(* IEC 61131-3 sources: ATCMcontrol_Engineering/src/COM/softing/fc/AddOns/Softing/4CPCTarget/Libs/ATCM_Communication, 12 files *)

(* ---- CONNECT.ST ---- *)
(*[[
    UserURL= "ATCM:CONNECT.htm"
]]*)

(* Communication Function Blocks, see IEC 1131-5
 * Implements the CONNECT communication function block
 *
*)

FUNCTION_BLOCK CONNECT      (* Connection management *)
VAR_INPUT
	EN_C    : BOOL := FALSE;   (* enable/startup connection *)
	PARTNER : COMM_PARTNER;    (* identifies communication partner and comm. deployment *)
END_VAR
VAR_OUTPUT
	VALID  : BOOL := FALSE;    (* connection is valid/established *)
	ERROR  : BOOL := FALSE;    (* new non-zero STATUS received *)
    STATUS : DINT := CFB_NoError;   (* last detected status *)
	ID     : COMM_CHANNEL;     (* established communication channel *)
END_VAR

VAR
    iType       : DINT;
    hChannel    : DINT;
    sParam      : WSTRING;
    bError   : BOOL;            (* true if error occured *)
    iNewStatus : DINT;          (* new status *)
    iFbState : DINT := 0;       (* state of function block:*)
                                (*  0: INIT
                                    1: IDLE
                                    2: CONNECTING
                                    3: CHECKING
                                    4: CONNECTED
                                    5: CLOSING
                                    6: CONCLUDING
                                    7: RETRY
                                    8: ABORT
                                    10: ERROR
                                *)
END_VAR

VAR_NATIVE
    static CommFBFactory g_commFBFact = new CommFBFactory();
    private CommFB comm = null;
    private int hChannel;
    private int iType;
    public void release()
    {
        if (comm != null)
        {
            CommFBFactory.removeCommFB(hChannel, iType);
            comm.closeConn();
            comm.release();
            comm = null;
        }
        super.release();
    }
END_VAR

VAR_NATIVE#movetop
import COM.softing.fc.CC.commFB.*;
END_VAR

(*
NATIVE
END_VAR
*)

(* Init local variables *)
hChannel := ID.hChannel;
iType := ID.iCommType;
bError := FALSE;
iNewStatus := CFB_NoError;

(* Init OutVars *)
ERROR := FALSE;

(* INIT funciton Block *)
IF iFbState = 0 THEN
    VALID := FALSE;
    STATUS := CFB_NoError;

    (* fast initialization => next fb state: idle *)
    iFbState := 1;
END_IF;

(* IDLE until new connect request *)
IF iFbState = 1 THEN
    IF EN_C THEN
        VALID := FALSE;
        ID.hChannel := -1;  (* not valid *)
        hChannel := -1;

        iType := PARTNER.iCommType;
        sParam := PARTNER.sParam;
        ID.iCommType := iType;
        ID.iTimeout := PARTNER.iTimeout;
        (* next state connecting *)
        iFbState := 2;
    ELSE
        (* Idle...*)
        RETURN;
    END_IF;
END_IF;

(* CONNECTING *)
IF iFbState = 2 THEN
    IF EN_C THEN
        (* Open connection *)
        NATIVE
        //if there is an old commFB, KILL IT NOW!
        if (comm != null)
        {
            CommFBFactory.removeCommFB(hChannel, iType);
            comm.closeConn();
            comm.release();
            comm = null;
        }
        // create new CommFB
        comm = CommFBFactory.createCommFB(iType = _itype.getInt());
        if (comm == null)
        {
            _berror.putBool(true);
            _inewstatus.putInt(-4); // CFB_ErrOutOfMemory
        }
        else
        {
            // open connection
            if (comm.openConn(_sparam.getString()))
            {
                hChannel = CommFBFactory.addCommFBToMap(comm);
                _hchannel.putInt(hChannel);
            }
            else
            {
                _berror.putBool(true);
                _inewstatus.putInt(comm.getConnStatus()); // CFB_...
                comm = null;
            }
        }
        END_NATIVE;

        IF bError THEN
            (* next state error *)
            iFbState := 10;
            GOTO error;
        ELSE
            (* next state checking *)
            iFbState := 3;
        END_IF;

    ELSE (* EN_C = FALSE *)
        (* Abort => next state idle *)
        iFbState := 1;
        RETURN;
    END_IF;
END_IF;

(* CHECKING *)
IF iFbState = 3 THEN
    NATIVE
    if (comm == null)
    {
        _berror.putBool(true);
        _inewstatus.putInt(7);  // CFB_ErrRemoteWrongState
        // next state error
        _ifbstate.putInt(10);
    }
    else if (!comm.checkConn())
    {
        _berror.putBool(true);
        _inewstatus.putInt(1);  // CFB_ErrLowLayer
        // next state abort
        _ifbstate.putInt(8);
    }
    END_NATIVE;

    IF bError = FALSE THEN
        ID.hChannel := hChannel;
        VALID := TRUE;
        (* next state connected *)
        iFbState := 4;
        (* wait for next cycle... *)
        RETURN;
    END_IF;
END_IF;

(* CONNECTED *)
IF iFbState = 4 THEN
    IF EN_C = FALSE THEN
        (* next state closing *)
        iFbState := 5;
    ELSE
        NATIVE
        if (comm == null)
            _berror.putBool(true);
        END_NATIVE;

        IF bError THEN
            iNewStatus := CFB_ErrRemoteWrongState;
            (* next state error *)
            iFbState := 10;
            GOTO error;
        ELSE
            (* check if connection is closed by the remote station *)
            NATIVE
            if (comm.isRemoteClosing())
            {
                // next state concluding
                _ifbstate.putInt(6);
                // wait for next cycle...
                return;
            }
            END_NATIVE;

            (* check if connection is still alive *)
            NATIVE
            if (!comm.checkConn())
            {
                _berror.putBool(true);
                _inewstatus.putInt(1); // CFB_ErrLowLayer
                // next state retry
                _ifbstate.putInt(7);
            }
            END_NATIVE;
        END_IF;
    END_IF;
END_IF;

(* CLOSING *)
IF iFbState = 5 THEN
    NATIVE
    if (comm != null)
    {
        CommFBFactory.removeCommFB(hChannel, iType);
        comm.closeConn();
        comm.release();
        comm = null;
    }
    END_NATIVE;

    VALID := FALSE;
    ID.hChannel := -1;
    (* next state idle *)
    iFbState := 1;
END_IF;

(* CONCLUDING *)
IF iFbState = 6 THEN
    NATIVE
    if (comm != null)
    {
        CommFBFactory.removeCommFB(hChannel, iType);
        comm.closeConn();
        comm.release();
        comm = null;
    }
    END_NATIVE;

    VALID := FALSE;
    ID.hChannel := -1;
    STATUS := CFB_ErrResetReceived;
    (* next state idle *)
    iFbState := 1;
END_IF;

(* RETRY *)
IF iFbState = 7 THEN
    NATIVE
    if (comm != null)
    {
        CommFBFactory.removeCommFB(hChannel, iType);
        comm.closeConn();
        comm.release();
        comm = null;
    }
    END_NATIVE;
    (* next state error *)
    iFbState := 10;
    GOTO error;
END_IF;

(* ABORT *)
IF iFbState = 8 THEN
    NATIVE
    if (comm != null)
    {
        CommFBFactory.removeCommFB(hChannel, iType);
        comm.closeConn();
        comm.release();
        comm = null;
    }
    END_NATIVE;
    (* next state error *)
    iFbState := 10;
    GOTO error;
END_IF;

(* ERROR *)
error:
IF iFbState = 10 THEN
    NATIVE
    if (comm != null)
    {
        CommFBFactory.removeCommFB(hChannel, iType);
        comm.closeConn();
        comm.release();
        comm = null;
    }
    END_NATIVE;

    VALID := FALSE;
    ERROR := TRUE;
    STATUS := iNewStatus;

    iFbState := 1;
    RETURN;
END_IF;

END_FUNCTION_BLOCK

(* ---- RCV.ST ---- *)
(*[[
]]*)

(* Communication Function Blocks, see IEC 1131-5
 * Implements the RCV communication function block
 *
*)

NATIVE
import COM.softing.fc.CC.commFB.*;
END_NATIVE

FUNCTION_BLOCK RCV      (* Interlocked control, responder*)
VAR_INPUT
    EN_R   : BOOL;          (* Enable to receive data *)
    RESP   : BOOL (*R_EDGE*);   (* Request to send response data *)
    ID     : COMM_CHANNEL;  (* Communication channel *)
    R_ID   : WSTRING;       (* Remote function block *)
    EXPECT : DINT;          (* non-IEC: number of bytes to receive *)
(*    SD_1   : ANY;*)           (* User data to send *)
(*    SD_m   : ANY; *)
END_VAR

VAR_OUTPUT
NDR    : BOOL;              (* New user data received *)
ERROR  : BOOL;              (* New non-zero STATUS received *)
STATUS : DINT;              (* Last detected status *)

RD_1   : WSTRING; (*ANY*)       (* Received user data *)
(*RD_n   : ANY;*)         (*  It is not required that m=n *)
END_VAR                 (*  either m, n, or both may be 0*)

    (* is not implemented yet !! *)
    ERROR := TRUE;
    STATUS := CFB_ErrNotImpl;

NATIVE
END_NATIVE;

END_FUNCTION_BLOCK

(* ---- SEND.ST ---- *)
(*[[
]]*)

(* Communication Function Blocks, see IEC 1131-5
 * Implements the SEND communication function block
 *
*)

NATIVE
import COM.softing.fc.CC.commFB.*;
END_NATIVE

FUNCTION_BLOCK SEND     (* Interlocked control, requester*)
VAR_INPUT
    REQ    : BOOL (*R_EDGE*);       (* Request to send with raising edge*)
    R      : BOOL (*R_EDGE*);       (* Reset local, remote function *)
    ID     : COMM_CHANNEL;      (* Communication channel *)
    R_ID   : WSTRING;           (* Remote function block *)
    SD_1   : WSTRING;  (*ANY*)  (* User data to send *)
END_VAR

VAR_OUTPUT
    NDR    : BOOL;          (* New user data received *)
    ERROR  : BOOL;        (* New non-zero STATUS received *)
    STATUS : DINT;        (* Last detected status *)
(*    RD_1   : ANY;*)         (* Received user data *)
END_VAR                 (*   either m, n, or both may be 0*)

    (* is not implemented yet !! *)
    ERROR := TRUE;
    STATUS := CFB_ErrNotImpl;

NATIVE
END_NATIVE;

END_FUNCTION_BLOCK

(* ---- SER_READ.ST ---- *)
(*[[
    UserURL= "ATCM:SER_READ.htm"
]]*)

(* Communication Function Blocks, see IEC 1131-5 for serial communication
 * Derived from the READ communication function block
 * differs in RD_LEN1, resp. RD_1 from READ in IEC 1131-5!
*)

FUNCTION_BLOCK SER_READ     (* Polled data acquisition *)
VAR_INPUT
    REQ      : BOOL R_EDGE := FALSE;    (* Request *)
    ID       : COMM_CHANNEL;    (* Communication channel *)
    RD_LEN_1 : DINT;            (* Min. length of the data to be received *)
    READ_ALL : BOOL := FALSE;   (* TRUE: all available data will be read, at least RD_LEN_1 *)
END_VAR

VAR_OUTPUT
    NDR    : BOOL;              (* New user data received *)
    ERROR  : BOOL;              (* New non-zero STATUS received *)
    STATUS : DINT;              (* Last detected status *)
    RD_1   : BYTE_STRING;       (* Received user data *)
END_VAR

VAR
    hChannel : DINT;
    iType    : DINT;
    bError   : BOOL;            (* true if error occured *)
    iNewStatus : DINT;          (* new status *)
    iFbState : DINT := 0;       (* state of function block:*)
                                (*  0: INIT
                                    1: IDLE
                                    2: WAITING
                                    3: CHECKING
                                    4: HAVE_DATA
                                    10: ERROR
                                *)
    timer    : TON;             (* timer for read timeout *)
    timer_IN : BOOL;
    timer_PT : TIME;
    bTimeout : BOOL;
END_VAR

VAR_NATIVE
    private CommFB comm;
END_VAR
VAR_NATIVE#movetop
import COM.softing.fc.CC.commFB.*;
import COM.softing.fc.CC.utility.*;
END_VAR

(* Init local variables*)
hChannel := ID.hChannel;
iType := ID.iCommType;
bError := FALSE;

(* Init OutVars *)
NDR := FALSE;
ERROR := FALSE;

(* INIT funciton Block *)
IF iFbState = 0 THEN
    STATUS := CFB_NoError;

    (* fast initialization => goto next state IDLE*)
    iFbState := 1;
END_IF;

(* get CommFB *)
NATIVE
    comm = CommFBFactory.lookUpCommFB(_hchannel.getInt(), _itype.getInt());
    if (comm == null)
    {
        _berror.putBool(true);
    }
END_NATIVE;
IF bError THEN
    iNewStatus := CFB_ErrInvalidCommChannel;
    iFbState := 10;
    GOTO error;
END_IF;

(* IDLE until new read request at raising edge of REQ input *)
IF iFbState = 1 THEN
    IF REQ THEN
        NATIVE
        // check if read is not active
        synchronized(comm) {
          if (comm.isReadActive())
            _berror.putBool(true);
          else
            comm.setReadActive(true);
        }
        END_NATIVE;

        IF bError THEN
            iNewStatus := CFB_ErrRemoteWrongState;
            iFbState := 10;
            GOTO error;
        END_IF;
        (* Start read request asynchronously *)
        (* reset timer *)
        bTimeout := FALSE;
        timer_IN := FALSE;
        timer_PT := DINT_TO_TIME(ID.iTimeout);
        timer(IN := timer_IN, PT := timer_PT);

        NATIVE
        // start read request
        if (!comm.readAsync(_rd_len_1, _read_all, (ByteString)_rd_1))
        {
            _berror.putBool(true);
            _inewstatus.putInt(comm.getReadStatus()); // CFB_...
            comm.setReadActive(false);
        }
        END_NATIVE;

        IF bError THEN
            iFBState := 10;
            GOTO error;
        END_IF;

        (* init new timer *)
        IF ID.iTimeout > 0 THEN
            timer_IN := TRUE;
        ELSE
            timer_IN := FALSE;
        END_IF;

        (* Next state WAITING *)
        iFbState := 2;

    ELSE
        (* Idle...*)
        RETURN;
    END_IF;
END_IF;

(* WAITING: wait for completion *)
IF iFbState = 2 THEN
    (* refresh timer *)
    timer(IN := timer_IN, PT := timer_PT);
    bTimeout := timer.Q;

    (* Wait for data *)
    NATIVE
    if (comm.hasReadCompleted())
    {
        // check status if error occured
        int iStat = comm.getReadStatus();
        if (iStat == 0)
        {
            // read finished : next state CHECKING
            _inewstatus.putInt(0);
            _ifbstate.putInt(3);
        }
        else
        {
            // error!
            _berror.putBool(true);
            _inewstatus.putInt(iStat); // CFB_...
            comm.setReadActive(false);
        }
    }
    else
    {
        // request pending!
        if (_btimeout.getBool())
        {
            // cancel read request
            comm.cancelReadRequest();
            _berror.putBool(true);
            comm.setReadActive(false);
        }
        else
        {
            // wait for next cycle...
            return;
        }
    }
    END_NATIVE;
    IF bError THEN
        IF bTimeout THEN
            iNewStatus := CFB_ErrTimeout;
        ELSE
            ; (* iNewStatus already set *)
        END_IF;
        iFBState := 10;
        GOTO error;
    END_IF;

END_IF;

(* CHECKING data type match *)
IF iFbState = 3 THEN
    NATIVE
    if (!comm.verifyData())
    {
        _berror.putBool(true);
        comm.setReadActive(false);
    }
    END_NATIVE;
    IF bError THEN
        iNewStatus := CFB_ErrTypeMismatch;
        iFBState := 10;
        GOTO error;
    ELSE
        (* next state: HAVE DATA *)
        iFBState := 4;
    END_IF;
END_IF;

(* HAVE DATA *)
IF iFbState = 4 THEN
    (* copy data to RD_1 *)
    NATIVE
    comm.depositData();
    comm.setReadActive(false);
    END_NATIVE;

    NDR := TRUE;
    ERROR := FALSE;
    STATUS := 0;

    (* next state: IDLE *)
    iFbState := 1;
    RETURN;
END_IF;

(* ERROR *)
error:
IF iFbState = 10 THEN
    NDR := FALSE;
    ERROR := TRUE;
    STATUS := iNewStatus;

    iFbState := 1;
    RETURN;
END_IF;

END_FUNCTION_BLOCK

(* ---- SER_WRITE.st ---- *)
(*[[
    UserURL= "ATCM:SER_WRITE.htm"
]]*)

(* Communication Function Blocks, see IEC 1131-5 for serial communication
 * Derived from the WRITE communication function block
 * differs in SD_1 from WRITE in IEC 1131-5!
*)

FUNCTION_BLOCK SER_WRITE            (* Parametric control *)
VAR_INPUT
    REQ    : BOOL R_EDGE := FALSE;  (* Request *)
    ID     : COMM_CHANNEL;          (* Communication channel *)
    SD_1   : BYTE_STRING ;          (* value of to be set *)
END_VAR

VAR_OUTPUT
    DONE   : BOOL;        (* Function performed *)
    ERROR  : BOOL;        (* New non-zero STATUS received *)
    STATUS : DINT;        (* Last detected status *)
END_VAR

VAR
    hChannel : DINT;
    iType    : DINT;
    bError   : BOOL;            (* true if error occured *)
    iNewStatus : DINT;          (* new status *)
    iFbState : DINT := 0;       (* state of function block:*)
                                (*  0: INIT
                                    1: IDLE
                                    2: WAITING
                                    4: HAVE_IT
                                    10: ERROR
                                *)
    timer    : TON;             (* timer for write timeout *)
    timer_IN : BOOL;
    timer_PT : TIME;
    bTimeout : BOOL;
END_VAR

VAR_NATIVE
    private CommFB comm;
END_VAR
VAR_NATIVE#movetop
import COM.softing.fc.CC.commFB.*;
import COM.softing.fc.CC.utility.*;
END_VAR

(* INIT local variables*)
hChannel := ID.hChannel;
iType := ID.iCommType;
bError := FALSE;

(* Init OutVars *)
DONE := FALSE;
ERROR := FALSE;

(* Init funciton Block *)
IF iFbState = 0 THEN
    STATUS := CFB_NoError;

    (* fast initialization => goto state IDLE *)
    iFbState := 1;
END_IF;

(* get CommFB *)
NATIVE
    comm = CommFBFactory.lookUpCommFB(_hchannel.getInt(), _itype.getInt());
    if (comm == null)
    {
        _berror.putBool(true);
    }
END_NATIVE;
IF bError THEN
    iNewStatus := CFB_ErrInvalidCommChannel;
    iFbState := 10;
    GOTO error;
END_IF;

(* IDLE until new write request at raising edge of REQ input *)
IF iFbState = 1 THEN
    IF REQ THEN
        NATIVE
        // check if write is not active
        synchronized(comm) {
          if (comm.isWriteActive())
            _berror.putBool(true);
          else
            comm.setWriteActive(true);
        }
        END_NATIVE;

        IF bError THEN
            iNewStatus := CFB_ErrRemoteWrongState;
            iFbState := 10;
            GOTO error;
        END_IF;

        (* Start write request asynchronously *)
        (* reset timer *)
        bTimeout := FALSE;
        timer_IN := FALSE;
        timer_PT := DINT_TO_TIME(ID.iTimeout);
        timer(IN := timer_IN, PT := timer_PT);

        NATIVE
        // source: locVars[2])
        if (!comm.writeAsync((ByteString)_sd_1))
        {
            _berror.putBool(true);
            _inewstatus.putInt(comm.getWriteStatus()); // CFB_...
            comm.setWriteActive(false);
        }
        END_NATIVE;

        IF bError THEN
            iFBState := 10;
            GOTO error;
        END_IF;

        (* init new timer *)
        IF ID.iTimeout > 0 THEN
            timer_IN := TRUE;
        ELSE
            timer_IN := FALSE;
        END_IF;

        (* Sext state WAITING *)
        iFbState := 2;

    ELSE
        (* Idle...*)
        RETURN;
    END_IF;
END_IF;

(* WAITING: wait for completion *)
IF iFbState = 2 THEN
    (* refresh timer *)
    timer(IN := timer_IN, PT := timer_PT);
    bTimeout := timer.Q;

    (* Wait for completion *)
    NATIVE
    if (comm.hasWriteCompleted())
    {
        // check status if error occured
        int iStat = comm.getWriteStatus();
        if (iStat == 0)
        {
            // write finished: next state HAVE IT
            _inewstatus.putInt(0);
            _ifbstate.putInt(4);
        }
        else
        {
            // error!
            _berror.putBool(true);
            _inewstatus.putInt(iStat); // CFB_...
            comm.setWriteActive(false);
        }
    }
    else
    {
        // request pending!
        if (_btimeout.getBool())
        {
            // cancel write request
            comm.cancelWriteRequest();
            _berror.putBool(true);
            comm.setWriteActive(false);
        }
        else
        {
            // wait for next cycle...
            return;
        }
    }
    END_NATIVE;
    IF bError THEN
        IF bTimeout THEN
            iNewStatus := CFB_ErrTimeout;
        ELSE
            ; (* iNewStatus already set *)
        END_IF;
        iFBState := 10;
        GOTO error;
    END_IF;

END_IF;

(* HAVE IT *)
IF iFbState = 4 THEN
    NATIVE
    comm.setWriteActive(false);
    END_NATIVE;
    DONE := TRUE;
    ERROR := FALSE;
    STATUS := 0;

    iFbState := 1;
    RETURN;
END_IF;

(* ERROR *)
error:
IF iFbState = 10 THEN
    DONE := FALSE;
    ERROR := TRUE;
    STATUS := iNewStatus;

    iFbState := 1;
    RETURN;
END_IF;

END_FUNCTION_BLOCK

(* ---- STATUS.ST ---- *)
(*[[
]]*)

(* Communication Function Blocks, see IEC 1131-5
 * Implements the STATUS communication function block
 *
*)

NATIVE
import COM.softing.fc.CC.commFB.*;
END_NATIVE

FUNCTION_BLOCK STATUS   (* Device verification - requester *)
VAR_INPUT
    REQ    : BOOL (*R_EDGE*);   (* Request *)
    ID     : COMM_CHANNEL;  (* Communication channel *)
END_VAR

VAR_OUTPUT
    NDR    : BOOL;        (* New user data received *)
    ERROR  : BOOL;        (* New non-zero STATUS received *)
    STATUS : DINT;        (* Last detected status *)
    PHYS   : DINT;        (* Physical status of remote *)
                          (*   communication partner   *)
    LOG    : DINT;        (* Logical status of remote *)
                          (*   communication partner   *)
    LOCAL  : ARRAY[0..7] OF WORD;  (* Local status of remote *)
END_VAR

    (* is not implemented yet !! *)
    ERROR := TRUE;
    STATUS := CFB_ErrNotImpl;
NATIVE
END_NATIVE;

END_FUNCTION_BLOCK

(* ---- UDP_CONNECT.st ---- *)
(*[[
    UserURL= "ATCM:UDP_CONNECT.htm"
]]*)

(*
 *  UDP datagram communication Function Blocks
 *  UDP_CONNECT allows to open and close a socket
 *  this FunctionBlock should be called only once, when the
 *  socket should be opened or closed
 *)

FUNCTION_BLOCK UDP_CONNECT

VAR_INPUT
    EN_C : BOOL;           (* true: open and connect the socket *)
                           (*   the field LocalPort of SOCKET_HANDLE has to be filled
                                with the local port number where the socket wants to
                                receive messages *)
                           (* false: close the socket *)
                           (* this FunctionBlock should be called only once, when the
                              socket should be opened or closed *)
END_VAR

VAR_IN_OUT
    SOCKET_HANDLE : UDP_SOCKET_HANDLE;  (* a structure that describes the socket *)
END_VAR

VAR_OUTPUT
    VALID        : BOOL;   (* shows if the socket is open or close *)
    ERROR        : BOOL;   (* error information *)
    ERROR_NR     : DINT;
    ERROR_STRING : WSTRING;
END_VAR

VAR
    portNr : DInt;
    bc     : BOOL;
END_VAR

VAR_NATIVE#movetop
    import COM.softing.fc.CC.commFB.*;
END_VAR

if EN_C then
    portNr := SOCKET_HANDLE.localPort;
    bc := SOCKET_HANDLE.broadcastSocket;
    native
        ((COM.softing.fc.CC.commFB.UDPSocketHandle)_socket_handle).open(
                                    _portnr.getInt(),
                                    _bc.getBool(),
                                    _error,
                                    _error_nr,
                                    _error_string);
    end_native;
    VALID := not Error;
else
    native
        ((COM.softing.fc.CC.commFB.UDPSocketHandle)_socket_handle).close(
                                    _error,
                                    _error_nr,
                                    _error_string);
    end_native;
    VALID := false;
end_if;
;
END_FUNCTION_BLOCK

(* ---- UDP_LOOKUP.st ---- *)
(*[[
    UserURL= "ATCM:UDP_LOOKUP.htm"
]]*)

(*
 *  UDP datagram communication Function Blocks
 *  UDP_LOOKUP looks up the ip-address (abc.def.ghi.jkl)
 *  for a hostname, this has to be used in UDP_USEND
 *  UDP_LOOKUP works asynchron because lookup can take a while
 *)

FUNCTION_BLOCK UDP_LOOKUP

VAR_INPUT
    EN_L          : Bool;               (* if ENABLE_Lookup = true, do lookup else
                                            do nothing *)
    HOST_NAME     : WString;            (* the name of the host to look up *)
END_VAR

VAR_IN_OUT
    SOCKET_HANDLE : UDP_SOCKET_HANDLE;  (* a handle to a opened socket *)
END_VAR

VAR_OUTPUT
    READY         : Bool;               (* shows that the lookup thread has finished *)
    HOST_ADDRESS  : WString;            (* if the lookup succeeded, the address of the host *)
    ERROR         : Bool;               (* error information if an error happened *)
    ERROR_NR      : DInt;
    ERROR_STRING  : WString;
END_VAR

VAR_NATIVE#movetop
    import COM.softing.fc.CC.commFB.*;
END_VAR

native
    ((COM.softing.fc.CC.commFB.UDPSocketHandle)_socket_handle).lookup(
                                    _en_l.getBool(),
                                    _host_name.getString(),
                                    _ready,
                                    _host_address,
                                    _error,
                                    _error_nr,
                                    _error_string);
end_native;

;
END_FUNCTION_BLOCK

(* ---- UDP_URCV.st ---- *)
(*[[
    UserURL= "ATCM:UDP_URCV.htm"
]]*)

(*
 *  UDP datagram communication Function Blocks
 *  UDP_URCV allows to receive a message from a partner
 *  through an open socket, URCV looks if there is a new msg
 *  available. If yes it returns the msg data, else NDR shows
 *  that no new msg is available
 *)

FUNCTION_BLOCK UDP_URCV

VAR_INPUT
    EN_R     : BOOL;            (* true: look for a new msg, false: do nothing *)
    DATA_LEN : DINT;            (* the maximum number of bytes that want to be received *)
                                (*  udp is a datagram based protocol, that means the
                                    data will be received in packets. If the available packet is
                                    longer than DATA_LEN, only DATA_LEN bytes will be returend,
                                    the rest is lost *)
END_VAR

VAR_IN_OUT
    SOCKET_HANDLE : UDP_SOCKET_HANDLE;  (* a structure that describes the socket *)
END_VAR

VAR_OUTPUT
    RD_1         : BYTE_STRING;  (* contains the msg data, if a new msg has been received *)
    PARTNER_ADDR : WSTRING;      (* the address and port of the communication partner *)
    PARTNER_PORT : DINT;         (*    that sent the received msg *)
    NDR          : BOOL;         (* shows if a new msg has been received *)
    ERROR        : BOOL;         (* error information *)
    ERROR_NR     : DINT;
    ERROR_STRING : WSTRING;
END_VAR

VAR_NATIVE#movetop
    import COM.softing.fc.CC.commFB.*;
END_VAR

if (EN_R) then
    native
        ((COM.softing.fc.CC.commFB.UDPSocketHandle)_socket_handle).receive(
                _data_len.getInt(),
                _rd_1,
                _partner_addr,
                _partner_port,
                _error,
                _error_nr,
                _error_string);
    end_native;
    if (RD_1.size>0) then
        NDR := true;
    else
        NDR := false;
    end_if;
end_if;
;
END_FUNCTION_BLOCK

(* ---- UDP_USEND.st ---- *)
(*[[
    UserURL= "ATCM:UDP_USEND.htm"
]]*)

(*
 *  UDP datagram communication Function Blocks
 *  UDP_USEND allows to send a message to a partner
 *  through an open socket
 *)

FUNCTION_BLOCK UDP_USEND

VAR_INPUT
    REQ          : BOOL;             (* true: send the msg, false: do nothing *)
    PARTNER_ADDR : WSTRING;          (* the host address of the communication partner *)
    PARTNER_PORT : DINT;             (* the port number where the comm. partner receives its msgs *)
    SD_1         : BYTE_STRING;      (* the data of the msg that will be sent *)
END_VAR

VAR_IN_OUT
    SOCKET_HANDLE : UDP_SOCKET_HANDLE; (* a structure that describes the socket *)
END_VAR

VAR_OUTPUT
    ERROR        : BOOL;             (* error information *)
    ERROR_NR     : DINT;
    ERROR_STRING : WSTRING;
END_VAR

VAR_NATIVE#movetop
    import COM.softing.fc.CC.commFB.*;
END_VAR

if (REQ) then
    native
        ((COM.softing.fc.CC.commFB.UDPSocketHandle)_socket_handle).send(
            _partner_addr.getString(),
            _partner_port.getInt(),
            _sd_1,
            _error,
            _error_nr,
            _error_string);
    end_native;
end_if;

END_FUNCTION_BLOCK

(* ---- USTATUS.ST ---- *)
(*[[
]]*)

(* Communication Function Blocks, see IEC 1131-5
 * Implements the USTATUS communication function block
 *
*)

NATIVE
import COM.softing.fc.CC.commFB.*;
END_NATIVE

FUNCTION_BLOCK USTATUS  (* Device verification - receiver *)
VAR_INPUT
    EN_R   : BOOL;        (* Enable to receive data *)
    ID     : COMM_CHANNEL;(* Communication channel *)
END_VAR

VAR_OUTPUT
    NDR    : BOOL;        (* New user data received *)
    ERROR  : BOOL;        (* New non-zero STATUS received *)
    STATUS : DINT;        (* Last detected status *)
    PHYS   : DINT;        (* Physical status of remote *)
                          (*   communication partner   *)
    LOG    : DINT;        (* Logical status of remote *)
                          (*   communication partner   *)
    LOCAL  : ARRAY[0..7] OF WORD; (* Local status of remote *)
                          (*   communication partner   *)
END_VAR

    (* is not implemented yet !! *)
    ERROR := TRUE;
    STATUS := CFB_ErrNotImpl;
NATIVE
END_NATIVE;

END_FUNCTION_BLOCK

(* ---- PrgTest.st ---- *)
(*[[
]]*)
PROGRAM PrgTest
var
    bstr     : byte_string;
    pos      : dint;
    valueIn  : wstring := "Umlaute: äöüßÄÖÜ andere Sachen: ´`°^";
    valueOut : wstring := "Umlaute: äöüßÄÖÜ andere Sachen: ´`°^";
    bError   : bool;
end_var

    pos := 0;
    COPY_WSTRING_TO_BYTE_STRING(valueIn, pos, bstr);

native
    try
    {
        byte byteString[] = ((COM.softing.fc.CC.utility.ByteString)_bstr).getByteString();
        java.io.FileOutputStream fi = new java.io.FileOutputStream("test.txt", false);
        fi.write(byteString);
        fi.close();
    }
    catch(java.io.IOException ioe)
    {
        _berror.putBool(true);
    }
end_native;

native
    try
    {
        byte byteString[] = ((COM.softing.fc.CC.utility.ByteString)_bstr).getByteString();
        java.io.FileInputStream fi = new java.io.FileInputStream("test.txt");
        fi.read(byteString);
        fi.close();
    }
    catch(java.io.IOException ioe)
    {
        _berror.putBool(true);
    }
end_native;

    pos := 0;
    valueOut := COPY_WSTRING_FROM_BYTE_STRING(bstr.size, pos, bstr);

END_PROGRAM
